(* IEC 61131-3 sources: codesys-to-astra/corpus/boiler-plc210/src/POUs/PRG_Fast, 2 files *)

(* ---- PRG_Fast.decl.st ---- *)
// Назначение: быстрые блокировки (задача FastTask, приоритет 0 у ОВЕН): авария горелки -> останов, сирена.
// Автор:      kr0nsch
// Версия:     0.1.0
// Документ:   corpus/boiler-plc210/README.md
PROGRAM PRG_Fast
VAR
END_VAR

(* ---- PRG_Fast.impl.st ---- *)
IF GVL_Hw.xBurner1Fault OR GVL_Hw.xBurner2Fault THEN
    GVL_Hmi.eState := E_BoilerState.Fault;
    GVL_Hw.xAlarmHorn := TRUE;
ELSE
    GVL_Hw.xAlarmHorn := FALSE;
END_IF
